Fanuc KAREL source: KD00004.KL

PROGRAM KD00004
%NOLOCKGROUP
%CRTDEVICE
VAR
  I: INTEGER
  J: INTEGER
  B: BOOLEAN
  R: REAL
  S: STRING[80]
BEGIN
  I = 1
END KD00004
